(* PLC project Unnamed, Unknown Unnamed 1 *)
(* stored: creationDateTime 2026-03-24T22:18:36, modificationDateTime 2026-05-19T17:14:10 *)

PROGRAM Exercise5
  VAR_INPUT
    Left_Hand : BOOL;
    Right_Hand : BOOL;
    Guard_Front : BOOL;
    Guard_Left : BOOL;
    Guard_Right : BOOL;
    E_Stop : BOOL;
    Mode_Switch : BOOL;
    Key_Switch : BOOL;
    Stroke_Sensor : BOOL;
    Both_Hands : BOOL;
  END_VAR
  VAR_OUTPUT
    Pressure_Pump : BOOL;
    Press_Ram_Full : BOOL;
    Press_Ram_Slow : BOOL;
    Safety_OK : BOOL;
    Fault_Light : BOOL;
    Pump_Run_Light : BOOL;
    Jam_Fault_Light : BOOL;
    Stabilization_Done : BOOL;
    Prev_Mode : BOOL;
    Mode_Changed : BOOL;
  END_VAR
  VAR
    TON0 : TON;
    TON1 : TON;
  END_VAR

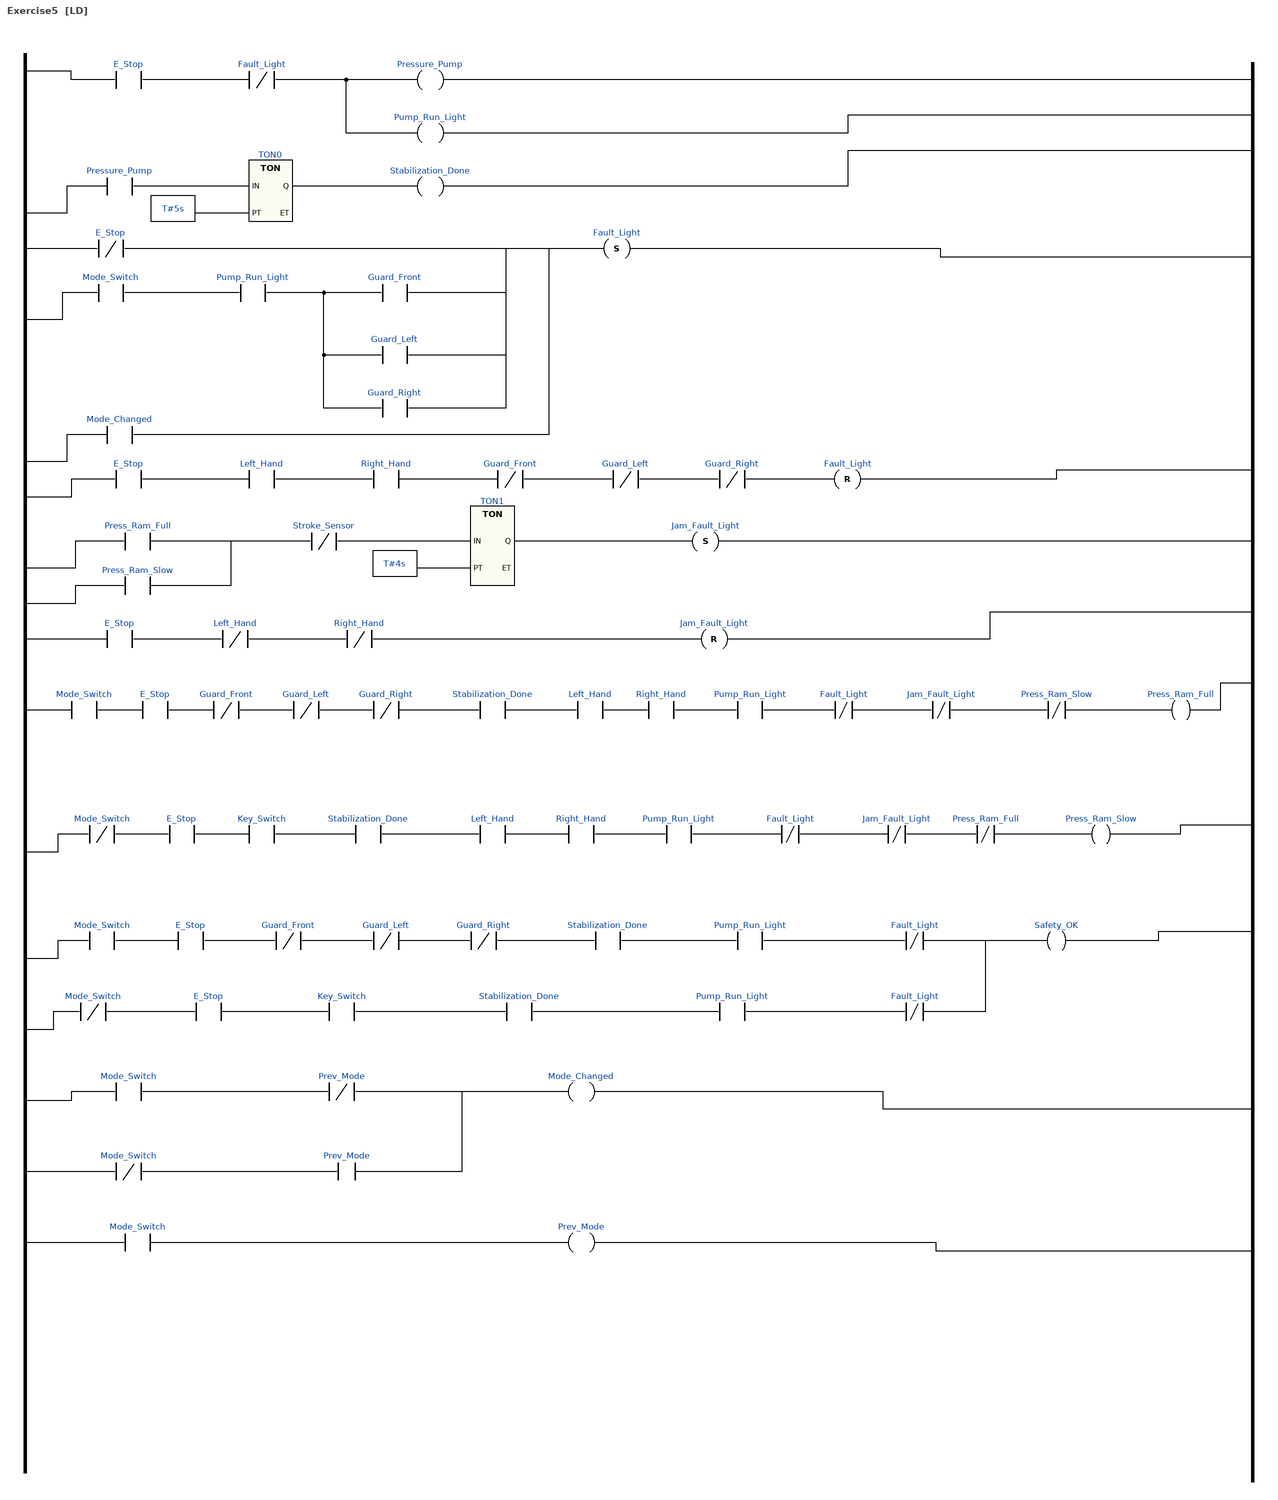
(* LD diagram, written out as Structured Text *)
Pressure_Pump := E_Stop AND NOT Fault_Light;
Pump_Run_Light := E_Stop AND NOT Fault_Light;
TON0(IN := Pressure_Pump, PT := T#5s);
Stabilization_Done := TON0.Q;
IF E_Stop AND Left_Hand AND Right_Hand AND NOT Guard_Front AND NOT Guard_Left AND NOT Guard_Right THEN Fault_Light := FALSE; END_IF;
IF NOT E_Stop OR Mode_Switch AND Pump_Run_Light AND Guard_Front OR Mode_Switch AND Pump_Run_Light AND Guard_Left OR Mode_Switch AND Pump_Run_Light AND Guard_Right OR Mode_Changed THEN Fault_Light := TRUE; END_IF;
TON1(IN := (Press_Ram_Full OR Press_Ram_Slow) AND NOT Stroke_Sensor, PT := T#4s);
IF TON1.Q THEN Jam_Fault_Light := TRUE; END_IF;
IF E_Stop AND NOT Left_Hand AND NOT Right_Hand THEN Jam_Fault_Light := FALSE; END_IF;
Press_Ram_Full := Mode_Switch AND E_Stop AND NOT Guard_Front AND NOT Guard_Left AND NOT Guard_Right AND Stabilization_Done AND Left_Hand AND Right_Hand AND Pump_Run_Light AND NOT Fault_Light AND NOT Jam_Fault_Light AND NOT Press_Ram_Slow;
Press_Ram_Slow := NOT Mode_Switch AND E_Stop AND Key_Switch AND Stabilization_Done AND Left_Hand AND Right_Hand AND Pump_Run_Light AND NOT Fault_Light AND NOT Jam_Fault_Light AND NOT Press_Ram_Full;
Safety_OK := Mode_Switch AND E_Stop AND NOT Guard_Front AND NOT Guard_Left AND NOT Guard_Right AND Stabilization_Done AND Pump_Run_Light AND NOT Fault_Light OR NOT Mode_Switch AND E_Stop AND Key_Switch AND Stabilization_Done AND Pump_Run_Light AND NOT Fault_Light;
Mode_Changed := Mode_Switch AND NOT Prev_Mode OR NOT Mode_Switch AND Prev_Mode;
Prev_Mode := Mode_Switch;
END_PROGRAM

CONFIGURATION Config0
  RESOURCE Res0 ON PLC
    TASK task0(INTERVAL := T#20ms, PRIORITY := 0);
    PROGRAM instance0 WITH task0 : Exercise5;
  END_RESOURCE
END_CONFIGURATION
